(* IEC 61131-3 sources: ironplc/integrations/vscode/src/screenshots/fixtures, 3 files *)

(* ---- invalid.st ---- *)
PROGRAM main
    VAR
        Button AT %IX1: BOOL;
        Buzzer AT %QX1: BOOL;
    END_VAR

    Buzzer := NOT Button;
    UndeclaredVar := 42;

END_PROGRAM

CONFIGURATION config
    RESOURCE res ON PLC
        TASK plc_task(INTERVAL := T#100ms, PRIORITY := 1);
        PROGRAM plc_task_instance WITH plc_task : main;
    END_RESOURCE
END_CONFIGURATION

(* ---- quickstart-helloworld.st ---- *)
PROGRAM main
   VAR
      Button : BOOL;
      Buzzer : BOOL;
   END_VAR

   Buzzer := NOT Button;

END_PROGRAM

(* ---- quickstart-timer.st ---- *)
PROGRAM main
   VAR
      Button : BOOL;
      Buzzer : BOOL;
      PulseTimer : TON;
   END_VAR

   PulseTimer(IN := NOT Button, PT := T#500ms);
   Buzzer := PulseTimer.Q;

END_PROGRAM

CONFIGURATION config
   RESOURCE res ON PLC
      TASK plc_task(INTERVAL := T#100ms, PRIORITY := 1);
      PROGRAM plc_task_instance WITH plc_task : main;
   END_RESOURCE
END_CONFIGURATION
